(*
SPDX-FileCopyrightText: c 2026 Oleksandr Tiutyk <trofimich@gmail.com>
SPDX-License-Identifier: MIT
License: https://opensource.org/license/mit
*)

(*!
<summary>Checks exact 255-unit and truncated 256-unit ANY text formatting.</summary>
<description>
Uses one task and stays at a stable address while assertions are bound to this instance.
</description>
*)

{attribute 'no_assign'}
{attribute 'no_explicit_call' := 'do not call this function block directly'}
FUNCTION_BLOCK WideStringLongFitFormattingTest EXTENDS TOF_Testing.SingleCycleTest
VAR_STAT
	{attribute 'hide'}
	_ClassName : STRING := __POUNAME();
END_VAR

(*!
<summary>Checks exact 255-unit and truncated 256-unit ANY text formatting.</summary>
<description>
Checks the retained code units, the U+2026 marker and the terminator directly in the returned buffer.
</description>
*)
METHOD PROTECTED ExecuteTest
VAR
	narrow : STRING(256);
	wide : WSTRING(256);
	wideData : POINTER TO WORD;
	result : WSTRING(255);
	resultData : POINTER TO WORD;
	i : INT;
END_VAR
wideData := ADR(wide);
resultData := ADR(result);

// SA0175: Fill STRING(256) with 256 ASCII bytes and terminate explicitly.
{analysis -175}
FOR i := 0 TO 255 DO
	narrow[i] := BYTE#16#61;
	wideData[i] := WORD#16#61;
END_FOR

narrow[256] := TO_BYTE(TOF_Core.UnsignedInt8.MIN_VALUE);
{analysis +175}
wideData[256] := TO_WORD(TOF_Core.UnsignedInt16.MIN_VALUE);

result := TOF_Core.WideStrings.AnyToStringFit255(value := narrow);
Assert.ThatBool(
	actual := TOF_Core.WideStrings.GetLength(value := result) = 255
		AND_THEN resultData[253] = WORD#16#61
		AND_THEN resultData[254] = WORD#16#2026
		AND_THEN resultData[255] = TO_WORD(TOF_Core.UnsignedInt16.MIN_VALUE),
	message := "A long STRING must retain 254 characters and append exactly U+2026"
).IsTrue();

result := TOF_Core.WideStrings.AnyToStringFit255(value := wide);
Assert.ThatBool(
	actual := TOF_Core.WideStrings.GetLength(value := result) = 255
		AND_THEN resultData[253] = WORD#16#61
		AND_THEN resultData[254] = WORD#16#2026
		AND_THEN resultData[255] = TO_WORD(TOF_Core.UnsignedInt16.MIN_VALUE),
	message := "A long WSTRING must retain 254 characters and append exactly U+2026"
).IsTrue();

// SA0175: Shorten the ASCII payload to exactly 255 bytes by moving its terminator.
{analysis -175}
narrow[255] := TO_BYTE(TOF_Core.UnsignedInt8.MIN_VALUE);
{analysis +175}
wideData[255] := TO_WORD(TOF_Core.UnsignedInt16.MIN_VALUE);
result := TOF_Core.WideStrings.AnyToStringFit255(value := narrow);
Assert.ThatBool(
	actual := TOF_Core.WideStrings.GetLength(value := result) = 255 AND_THEN resultData[254] = WORD#16#61,
	message := "An exact-fit STRING must keep its final character"
).IsTrue();
result := TOF_Core.WideStrings.AnyToStringFit255(value := wide);
Assert.ThatBool(
	actual := TOF_Core.WideStrings.GetLength(value := result) = 255 AND_THEN resultData[254] = WORD#16#61,
	message := "An exact-fit WSTRING must keep its final character"
).IsTrue();
END_METHOD

//! <summary>Borrows the concrete class name. Callers must not modify it.</summary>
{attribute 'monitoring' := 'call'}
PROPERTY ClassName : REFERENCE TO STRING
GET
ClassName REF= _ClassName;
END_GET
END_PROPERTY

//! <summary>Borrows the compiler-initialized namespace name. Callers must not modify it.</summary>
{attribute 'monitoring' := 'call'}
PROPERTY NamespaceName : REFERENCE TO STRING
GET
NamespaceName REF= CurrentNamespace.Name;
END_GET
END_PROPERTY

//! <summary>Reports the concrete instance size in bytes.</summary>
{attribute 'monitoring' := 'call'}
PROPERTY SelfSize : ULINT
GET
SelfSize := XSIZEOF(THIS^);
END_GET
END_PROPERTY

END_FUNCTION_BLOCK

(* stored: Version 1.1.0.1
   POU WideStringLongFitFormattingTest: Id {a026e757-e771-44ce-971b-36082a76d984}, SpecialFunc None
   Method ExecuteTest: Id {9f2f7f1a-56ea-4a64-9a7d-7620baccbe0e}
   Property ClassName: Id {ad8bb01b-79f2-41e0-9b16-488c6e3da590}
   Get Get: Id {0b9ab670-c7e4-47f6-983c-26ed6da8e0a2}
   Property NamespaceName: Id {60039231-a61b-4cd2-85a5-d205081f383a}
   Get Get: Id {e0fab7de-61ad-41aa-b541-3e4d711e3f28}
   Property SelfSize: Id {96b1369e-63e9-43e4-86b6-c032f1bc2bb8}
   Get Get: Id {05970a0d-d352-46b6-a8f1-4aef55e296ac} *)
